(* IEC 61131-3 sources: volt/packages/volt-lsp-iec/test-corpus/awa-palletizer/Device/Plc Logic/Application/Library Manager/Standard, 22 files *)

(* ---- CONCAT.pou ---- *)
FUNCTION CONCAT : STRING(255)
VAR_INPUT
	STR1 : STRING(255);
	STR2 : STRING(255);
END_VAR
END_FUNCTION

(* ---- DELETE.pou ---- *)
FUNCTION DELETE : STRING(255)
VAR_INPUT
	STR : STRING(255);
	LEN : INT;
	POS : INT;
END_VAR
END_FUNCTION

(* ---- FIND.pou ---- *)
FUNCTION FIND : INT
VAR_INPUT
	STR1 : STRING(255);
	STR2 : STRING(255);
END_VAR
END_FUNCTION

(* ---- INSERT.pou ---- *)
FUNCTION INSERT : STRING(255)
VAR_INPUT
	STR1 : STRING(255);
	STR2 : STRING(255);
	POS : INT;
END_VAR
END_FUNCTION

(* ---- LEFT.pou ---- *)
FUNCTION LEFT : STRING(255)
VAR_INPUT
	STR : STRING(255);
	SIZE : INT;
END_VAR
END_FUNCTION

(* ---- LEN.pou ---- *)
FUNCTION LEN : INT
VAR_INPUT
	STR : STRING(255);
END_VAR
END_FUNCTION

(* ---- LEN_INTERNAL.pou ---- *)
FUNCTION LEN_INTERNAL : UINT
VAR_IN_OUT
	STR : STRING(255);
END_VAR
END_FUNCTION

(* ---- MEMCOPY_INTERNAL.pou ---- *)
FUNCTION MEMCOPY_INTERNAL : POINTER TO BYTE
VAR_INPUT
	PDEST : POINTER TO BYTE;
	PSRC : POINTER TO BYTE;
	DWSIZE : DWORD;
END_VAR
END_FUNCTION

(* ---- MID.pou ---- *)
FUNCTION MID : STRING(255)
VAR_INPUT
	STR : STRING(255);
	LEN : INT;
	POS : INT;
END_VAR
END_FUNCTION

(* ---- REPLACE.pou ---- *)
FUNCTION REPLACE : STRING(255)
VAR_INPUT
	STR1 : STRING(255);
	STR2 : STRING(255);
	L : INT;
	P : INT;
END_VAR
END_FUNCTION

(* ---- RIGHT.pou ---- *)
FUNCTION RIGHT : STRING(255)
VAR_INPUT
	STR : STRING(255);
	SIZE : INT;
END_VAR
END_FUNCTION

(* ---- CTD.pou ---- *)
FUNCTION_BLOCK CTD
VAR_INPUT
	CD : BOOL;
	LOAD : BOOL;
	PV : WORD;
END_VAR
VAR_OUTPUT
	Q : BOOL;
	CV : WORD;
END_VAR
VAR
	M : BOOL;
END_VAR
END_FUNCTION_BLOCK

(* ---- CTU.pou ---- *)
FUNCTION_BLOCK CTU
VAR_INPUT
	CU : BOOL;
	RESET : BOOL;
	PV : WORD;
END_VAR
VAR_OUTPUT
	Q : BOOL;
	CV : WORD;
END_VAR
VAR
	M : BOOL;
END_VAR
END_FUNCTION_BLOCK

(* ---- CTUD.pou ---- *)
FUNCTION_BLOCK CTUD
VAR_INPUT
	CU : BOOL;
	CD : BOOL;
	RESET : BOOL;
	LOAD : BOOL;
	PV : WORD;
END_VAR
VAR_OUTPUT
	QU : BOOL;
	QD : BOOL;
	CV : WORD;
END_VAR
VAR
	MU : BOOL;
	MD : BOOL;
	RU : BOOL;
	RD : BOOL;
END_VAR
END_FUNCTION_BLOCK

(* ---- F_TRIG.pou ---- *)
FUNCTION_BLOCK F_TRIG
VAR_INPUT
	CLK : BOOL;
END_VAR
VAR_OUTPUT
	Q : BOOL;
END_VAR
VAR
	M : BOOL := TRUE;
END_VAR
END_FUNCTION_BLOCK

(* ---- R_TRIG.pou ---- *)
FUNCTION_BLOCK R_TRIG
VAR_INPUT
	CLK : BOOL;
END_VAR
VAR_OUTPUT
	Q : BOOL;
END_VAR
VAR
	M : BOOL;
END_VAR
END_FUNCTION_BLOCK

(* ---- RS.pou ---- *)
FUNCTION_BLOCK RS
VAR_INPUT
	SET : BOOL;
	RESET1 : BOOL;
END_VAR
VAR_OUTPUT
	Q1 : BOOL;
END_VAR
END_FUNCTION_BLOCK

(* ---- RTC.pou ---- *)
FUNCTION_BLOCK RTC
VAR_INPUT
	EN : BOOL;
	PDT : DATE_AND_TIME;
END_VAR
VAR_OUTPUT
	Q : BOOL;
	CDT : DATE_AND_TIME;
END_VAR
VAR
	M : BOOL;
	DIFFTIME : TIME;
	LASTTIME : TIME := TIME#0ms;
	TIMEOFFSET : TIME := TIME#0ms;
	CURTIME : TIME;
END_VAR
END_FUNCTION_BLOCK

(* ---- SR.pou ---- *)
FUNCTION_BLOCK SR
VAR_INPUT
	SET1 : BOOL;
	RESET : BOOL;
END_VAR
VAR_OUTPUT
	Q1 : BOOL;
END_VAR
END_FUNCTION_BLOCK

(* ---- TOF.pou ---- *)
FUNCTION_BLOCK TOF
VAR_INPUT
	IN : BOOL;
	PT : TIME;
END_VAR
VAR_OUTPUT
	Q : BOOL;
	ET : TIME;
END_VAR
VAR
	M : BOOL;
	STARTTIME : TIME;
END_VAR
END_FUNCTION_BLOCK

(* ---- TON.pou ---- *)
FUNCTION_BLOCK TON
VAR_INPUT
	IN : BOOL;
	PT : TIME;
END_VAR
VAR_OUTPUT
	Q : BOOL;
	ET : TIME;
END_VAR
VAR
	M : BOOL;
	STARTTIME : TIME;
END_VAR
END_FUNCTION_BLOCK

(* ---- TP.pou ---- *)
FUNCTION_BLOCK TP
VAR_INPUT
	IN : BOOL;
	PT : TIME;
END_VAR
VAR_OUTPUT
	Q : BOOL;
	ET : TIME;
END_VAR
VAR
	STARTTIME : TIME;
END_VAR
END_FUNCTION_BLOCK
